// État d'un OF dans la table du PLC (docs/05 § 5.6)
{attribute 'qualified_only'}
{attribute 'strict'}
TYPE E_OrderState :
(
    Free := 0,
    Active := 1,
    Suspended := 2,
    Done := 3
) USINT;
END_TYPE

(* stored: Version 1.1.0.1, ProductVersion 3.1.4024.12
   DUT E_OrderState: Id {274ec2ff-95e1-588f-ad6f-79a261ccec6e} *)
